(* IEC 61131-3 sources: plc-process-lib/src/POUs/Util/F_IsFinite, 2 files *)

(* ---- F_IsFinite.decl.st ---- *)
// Назначение: TRUE, если REAL — конечное правдоподобное число. FALSE для NaN и ±Inf
//             (все биты экспоненты = 1, проверка по битам через U_RealBits — не зависит от
//             оптимизатора) и для |rIn| > REAL_SANE_MAX (мусор: перепутан порядок слов Modbus).
// Автор:      kr0nsch
// Версия:     0.1.0
// Документ:   docs/fb/Functions.md
FUNCTION F_IsFinite : BOOL
VAR_INPUT
    rIn : REAL;            // проверяемое значение
END_VAR
VAR
    uBits : U_RealBits;    // биты значения
END_VAR

(* ---- F_IsFinite.impl.st ---- *)
uBits.rValue := rIn;
IF (uBits.dwValue AND GVL_Const.REAL_EXP_MASK) = GVL_Const.REAL_EXP_MASK THEN
    // экспонента из одних единиц: NaN, +Inf или -Inf
    F_IsFinite := FALSE;
ELSE
    // конечное число: ABS не дойдёт до NaN
    F_IsFinite := ABS(rIn) <= GVL_Const.REAL_SANE_MAX;
END_IF
